Staubli VAL3: Lab2B.dtx


